FUNCTION_BLOCK TestCtrl (* Basic Function Block Type *)
  (* Standard: 61499-2 *)
  (* Version 0.0, 7/2/2026, Template *)
  PACKAGE Main;
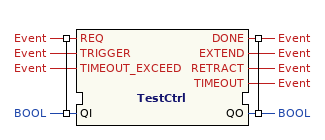
  EVENT_INPUT
    REQ WITH QI; (* Normal Execution Request *)
    TRIGGER;
    TIMEOUT_EXCEED;
  END_EVENT
  EVENT_OUTPUT
    DONE WITH QO;
    EXTEND;
    RETRACT;
    TIMEOUT;
  END_EVENT
  VAR_INPUT
    QI : BOOL; (* Input event qualifier *)
  END_VAR
  VAR_OUTPUT
    QO : BOOL; (* Output event qualifier *)
  END_VAR
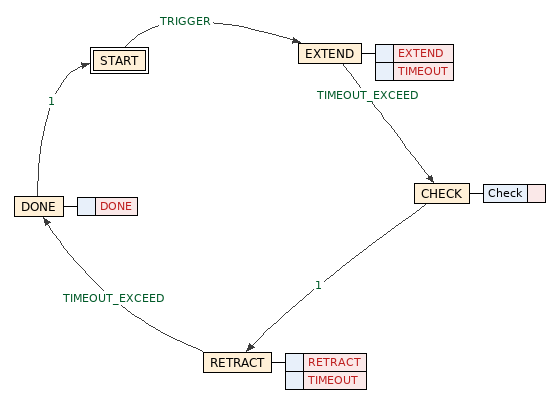
  EC_STATES
    START; (* Initial State *)
    EXTEND : -> EXTEND, -> TIMEOUT;
    CHECK : Check;
    RETRACT : -> RETRACT, -> TIMEOUT;
    DONE : -> DONE;
  END_STATES
  EC_TRANSITIONS
    DONE TO START := 1;
    START TO EXTEND := TRIGGER;
    EXTEND TO CHECK := TIMEOUT_EXCEED;
    RETRACT TO DONE := TIMEOUT_EXCEED;
    CHECK TO RETRACT := 1;
  END_TRANSITIONS
  ALGORITHM INIT IN ST: (* Initialization algorithm *)
;
  END_ALGORITHM
  ALGORITHM REQ IN ST: (* Normally executed algorithm *)
;
  END_ALGORITHM
  ALGORITHM Check IN ST:
QO:=QI;
  END_ALGORITHM
END_FUNCTION_BLOCK
